Staubli VAL3: CurrentTool.dtx

public num nItem
public tool tValue = {fatherId=flange[0]}
public string sName
public num nItemM
